{attribute 'strict'}
{attribute 'to_string'}
TYPE E_YARD_CHECK :
(
  NULL,

  POINTER_CTRL_INVALID                := 9000,
  POINTER_STATE_INVALID,
  REFERENCE_INSTANCE_CONTROL_INVALID,
  REFERENCE_INSTANCE_STATE_INVALID,

	POINTER_TRANSPORT_CTRL_INVALID      := 9100,
	POINTER_TRANSPORT_STATE_INVALID     := 9200,
	POINTER_COLLECTOR_ITF_INVALID       := 9300,
  REFERENCE_TICKET_LIST_ITF_INVALID   := 9400,

  CHECK_DONE := 10000

)UINT;
END_TYPE

(* stored: Version 1.1.0.1
   DUT E_YARD_CHECK: Id {133628a9-edd6-478b-89b2-3c6005d26235} *)
